Omron CX-Programmer project OmronTeachingExample (CX-Programmer 9.73)

# PLC ExamplePLC: CP1H XA

## Program Main (cyclic task 0)

### Section Section1

### Section Signed32_Constants

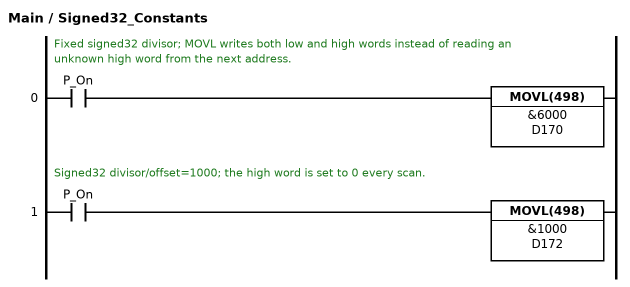
; rung 0: Fixed signed32 divisor; MOVL writes both low and high words instead of reading an unknown high word from the next address.
LD P_On
MOVL(498) &6000 D170
; rung 1: Signed32 divisor/offset=1000; the high word is set to 0 every scan.
LD P_On
MOVL(498) &1000 D172

### Section Analog_Validity

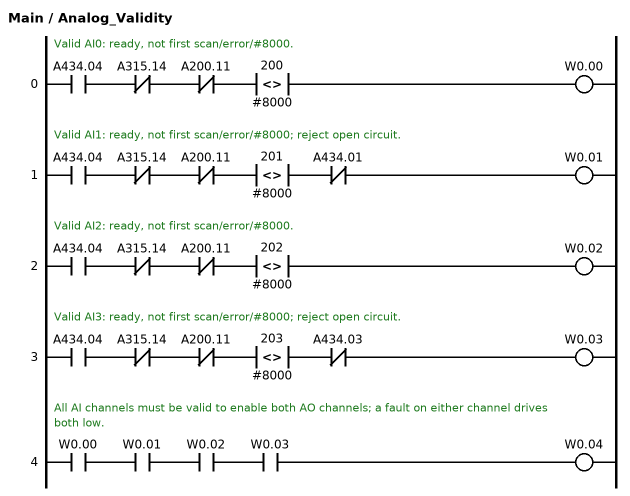
; rung 0: Valid AI0: ready, not first scan/error/#8000.
LD A434.04
ANDNOT A315.14
ANDNOT A200.11
AND<>(305) 200 #8000
OUT W0.00
; rung 1: Valid AI1: ready, not first scan/error/#8000; reject open circuit.
LD A434.04
ANDNOT A315.14
ANDNOT A200.11
AND<>(305) 201 #8000
ANDNOT A434.01
OUT W0.01
; rung 2: Valid AI2: ready, not first scan/error/#8000.
LD A434.04
ANDNOT A315.14
ANDNOT A200.11
AND<>(305) 202 #8000
OUT W0.02
; rung 3: Valid AI3: ready, not first scan/error/#8000; reject open circuit.
LD A434.04
ANDNOT A315.14
ANDNOT A200.11
AND<>(305) 203 #8000
ANDNOT A434.03
OUT W0.03
; rung 4: All AI channels must be valid to enable both AO channels; a fault on either channel drives both low.
LD W0.00
AND W0.01
AND W0.02
AND W0.03
OUT W0.04

### Section HMI_Input_Publication

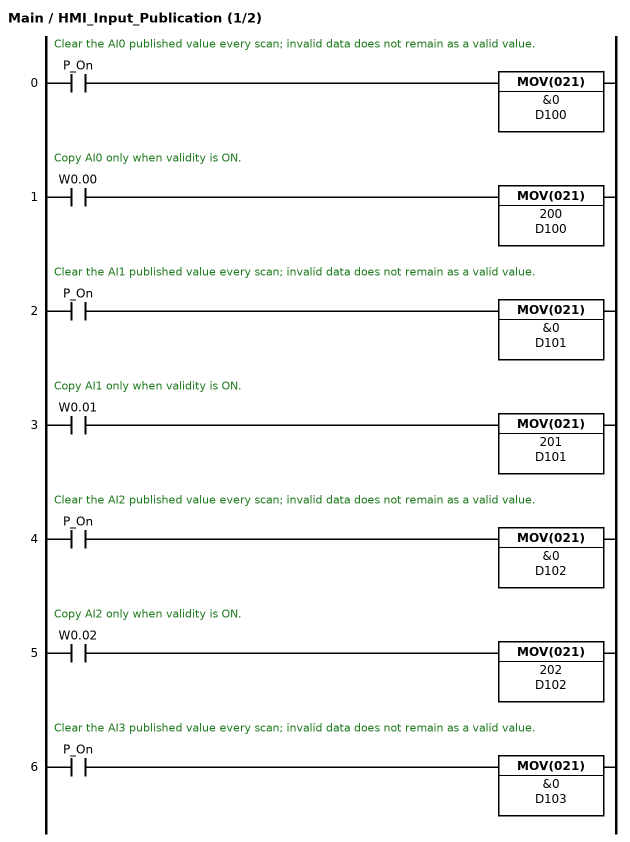
; rung 0: Clear the AI0 published value every scan; invalid data does not remain as a valid value.
LD P_On
MOV(021) &0 D100
; rung 1: Copy AI0 only when validity is ON.
LD W0.00
MOV(021) 200 D100
; rung 2: Clear the AI1 published value every scan; invalid data does not remain as a valid value.
LD P_On
MOV(021) &0 D101
; rung 3: Copy AI1 only when validity is ON.
LD W0.01
MOV(021) 201 D101
; rung 4: Clear the AI2 published value every scan; invalid data does not remain as a valid value.
LD P_On
MOV(021) &0 D102
; rung 5: Copy AI2 only when validity is ON.
LD W0.02
MOV(021) 202 D102
; rung 6: Clear the AI3 published value every scan; invalid data does not remain as a valid value.
LD P_On
MOV(021) &0 D103

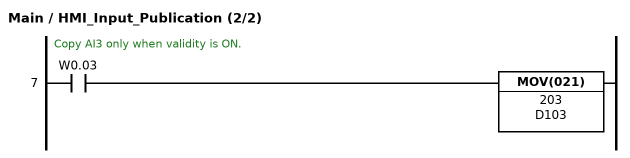
; rung 7: Copy AI3 only when validity is ON.
LD W0.03
MOV(021) 203 D103

### Section Math_Defaults_Each_Scan

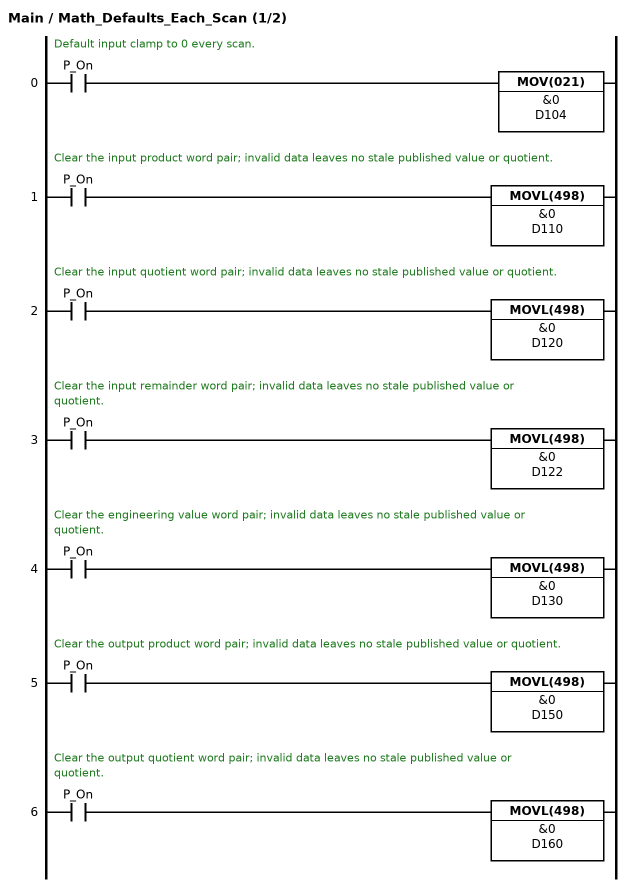
; rung 0: Default input clamp to 0 every scan.
LD P_On
MOV(021) &0 D104
; rung 1: Clear the input product word pair; invalid data leaves no stale published value or quotient.
LD P_On
MOVL(498) &0 D110
; rung 2: Clear the input quotient word pair; invalid data leaves no stale published value or quotient.
LD P_On
MOVL(498) &0 D120
; rung 3: Clear the input remainder word pair; invalid data leaves no stale published value or quotient.
LD P_On
MOVL(498) &0 D122
; rung 4: Clear the engineering value word pair; invalid data leaves no stale published value or quotient.
LD P_On
MOVL(498) &0 D130
; rung 5: Clear the output product word pair; invalid data leaves no stale published value or quotient.
LD P_On
MOVL(498) &0 D150
; rung 6: Clear the output quotient word pair; invalid data leaves no stale published value or quotient.
LD P_On
MOVL(498) &0 D160

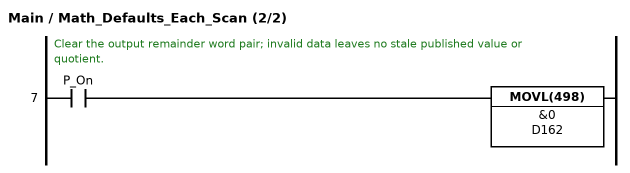
; rung 7: Clear the output remainder word pair; invalid data leaves no stale published value or quotient.
LD P_On
MOVL(498) &0 D162

### Section Signed32_Input_Scaling

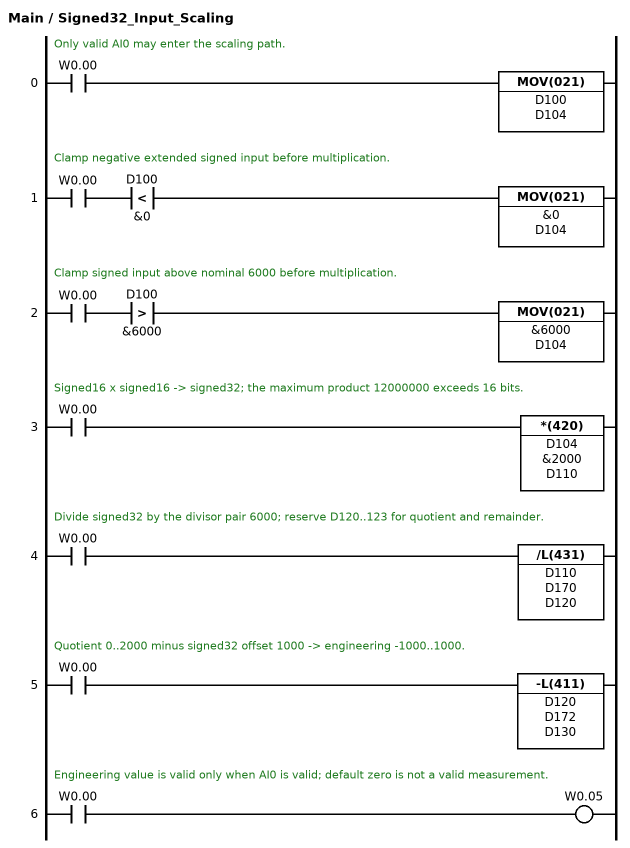
; rung 0: Only valid AI0 may enter the scaling path.
LD W0.00
MOV(021) D100 D104
; rung 1: Clamp negative extended signed input before multiplication.
LD W0.00
AND<S(312) D100 &0
MOV(021) &0 D104
; rung 2: Clamp signed input above nominal 6000 before multiplication.
LD W0.00
AND>S(322) D100 &6000
MOV(021) &6000 D104
; rung 3: Signed16 x signed16 -> signed32; the maximum product 12000000 exceeds 16 bits.
LD W0.00
*(420) D104 &2000 D110
; rung 4: Divide signed32 by the divisor pair 6000; reserve D120..123 for quotient and remainder.
LD W0.00
/L(431) D110 D170 D120
; rung 5: Quotient 0..2000 minus signed32 offset 1000 -> engineering -1000..1000.
LD W0.00
-L(411) D120 D172 D130
; rung 6: Engineering value is valid only when AI0 is valid; default zero is not a valid measurement.
LD W0.00
OUT W0.05

### Section Output_Scaling_And_Final_Writer

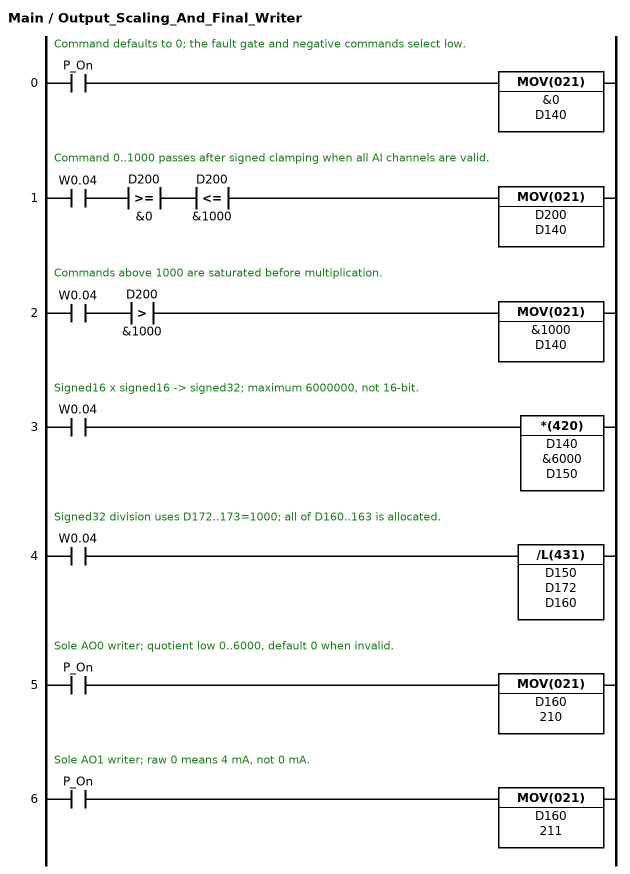
; rung 0: Command defaults to 0; the fault gate and negative commands select low.
LD P_On
MOV(021) &0 D140
; rung 1: Command 0..1000 passes after signed clamping when all AI channels are valid.
LD W0.04
AND>=S(327) D200 &0
AND<=S(317) D200 &1000
MOV(021) D200 D140
; rung 2: Commands above 1000 are saturated before multiplication.
LD W0.04
AND>S(322) D200 &1000
MOV(021) &1000 D140
; rung 3: Signed16 x signed16 -> signed32; maximum 6000000, not 16-bit.
LD W0.04
*(420) D140 &6000 D150
; rung 4: Signed32 division uses D172..173=1000; all of D160..163 is allocated.
LD W0.04
/L(431) D150 D172 D160
; rung 5: Sole AO0 writer; quotient low 0..6000, default 0 when invalid.
LD P_On
MOV(021) D160 210
; rung 6: Sole AO1 writer; raw 0 means 4 mA, not 0 mA.
LD P_On
MOV(021) D160 211

### Section END
; rung 0
END(001)